RESOURCE_TYPE TestResource (* Resource type with a basic FB *)
  (* Standard: 61499-1; Description: Copyright (c) 2026 Martin Erich Jobst This program and the accompanying materials are made available under the terms of the Eclipse Public License 2.0 which is available at https://www.eclipse.org/legal/epl-2.0/ SPDX-License-Identifier: EPL-2.0 *)
  (* Version 1.0, 2026-10-23, Martin Jobst *)
  {SET_ATTRIBUTE(IntegerAttribute, 14)}
  VAR_INPUT
    RESOURCE_ID : DINT := DINT#2;
  END_VAR
  FBS
    Processor : fixture::basic::BasicTest(DI1 := DINT#3); {SET_ATTRIBUTE(IntegerAttribute, 13)}
    Controller : CompositeTest;
  END_FBS
  SUBAPPS
    TypedSubApp : TestSubApp(DI1 := DINT#8); (* Configured typed subapplication *)
  END_SUBAPPS
END_RESOURCE_TYPE
